(* IEC 61131-3 sources: trust-platform/examples/OSCAT/cleanroom_pressure_strategy_composite/oop/src, 3 files *)

(* ---- Main.st ---- *)
(* Pattern role: IRoomNode is the contract boundary for the Strategy and Composite example. *)
INTERFACE IRoomNode
    PROPERTY ChildCount : INT
    GET
    END_GET
    END_PROPERTY
    PROPERTY PressureError : REAL
    GET
    END_GET
    END_PROPERTY
    PROPERTY AlarmCount : INT
    GET
    END_GET
    END_PROPERTY
    METHOD GetChild : IRoomNode
    VAR_INPUT
        Index : INT;
    END_VAR
    END_METHOD
END_INTERFACE

(* Pattern role: IPressureStrategy is the contract boundary for the Strategy and Composite example. *)
INTERFACE IPressureStrategy
    PROPERTY ModeId : INT
    GET
    END_GET
    END_PROPERTY
    METHOD TargetPressure : REAL
    VAR_INPUT
        BasePressurePa : REAL;
    END_VAR
    END_METHOD
END_INTERFACE

(* Pattern role: NormalPressureStrategy is a concrete implementation in the Strategy and Composite example. *)
FUNCTION_BLOCK NormalPressureStrategy IMPLEMENTS IPressureStrategy
METHOD PUBLIC TargetPressure : REAL
VAR_INPUT
    BasePressurePa : REAL;
END_VAR
TargetPressure := BasePressurePa;
END_METHOD
PUBLIC PROPERTY ModeId : INT
GET
    ModeId := INT#1;
END_GET
END_PROPERTY
END_FUNCTION_BLOCK

(* Pattern role: CleaningPressureStrategy is a concrete implementation in the Strategy and Composite example. *)
FUNCTION_BLOCK CleaningPressureStrategy IMPLEMENTS IPressureStrategy
METHOD PUBLIC TargetPressure : REAL
VAR_INPUT
    BasePressurePa : REAL;
END_VAR
TargetPressure := BasePressurePa + REAL#5.0;
END_METHOD
PUBLIC PROPERTY ModeId : INT
GET
    ModeId := INT#2;
END_GET
END_PROPERTY
END_FUNCTION_BLOCK

(* Pattern role: EmergencyPressureStrategy is a concrete implementation in the Strategy and Composite example. *)
FUNCTION_BLOCK EmergencyPressureStrategy IMPLEMENTS IPressureStrategy
METHOD PUBLIC TargetPressure : REAL
VAR_INPUT
    BasePressurePa : REAL;
END_VAR
TargetPressure := REAL#0.0;
END_METHOD
PUBLIC PROPERTY ModeId : INT
GET
    ModeId := INT#3;
END_GET
END_PROPERTY
END_FUNCTION_BLOCK

(* Pattern role: RoomNode is a concrete implementation in the Strategy and Composite example. *)
FUNCTION_BLOCK RoomNode IMPLEMENTS IRoomNode
VAR
    ErrorValue : REAL;
    AlarmValue : BOOL;
END_VAR
METHOD PUBLIC UpdateRoom
VAR_INPUT
    ActualPressurePa : REAL;
    TargetPressurePa : REAL;
    DoorOpen : BOOL;
END_VAR
ErrorValue := TargetPressurePa - ActualPressurePa;
AlarmValue := (ABS(ErrorValue) > REAL#10.0) OR DoorOpen;
END_METHOD
METHOD PUBLIC GetChild : IRoomNode
VAR_INPUT
    Index : INT;
END_VAR
GetChild := THIS;
END_METHOD
PUBLIC PROPERTY ChildCount : INT
GET
    ChildCount := INT#0;
END_GET
END_PROPERTY
PUBLIC PROPERTY PressureError : REAL
GET
    PressureError := ErrorValue;
END_GET
END_PROPERTY
PUBLIC PROPERTY AlarmCount : INT
GET
    IF AlarmValue THEN AlarmCount := INT#1; ELSE AlarmCount := INT#0; END_IF;
END_GET
END_PROPERTY
END_FUNCTION_BLOCK

(* Pattern role: RoomSuite is a concrete implementation in the Strategy and Composite example. *)
FUNCTION_BLOCK RoomSuite IMPLEMENTS IRoomNode
VAR
    Room1 : RoomNode;
    Room2 : RoomNode;
END_VAR
METHOD PUBLIC UpdateSuite
VAR_INPUT
    Room1Pressure : REAL;
    Room2Pressure : REAL;
    TargetPressure : REAL;
    DoorOpen : BOOL;
END_VAR
Room1.UpdateRoom(ActualPressurePa := Room1Pressure, TargetPressurePa := TargetPressure, DoorOpen := DoorOpen);
Room2.UpdateRoom(ActualPressurePa := Room2Pressure, TargetPressurePa := TargetPressure - REAL#5.0, DoorOpen := FALSE);
END_METHOD
METHOD PUBLIC GetChild : IRoomNode
VAR_INPUT
    Index : INT;
END_VAR
IF Index = INT#1 THEN GetChild := Room1; ELSE GetChild := Room2; END_IF;
END_METHOD
PUBLIC PROPERTY ChildCount : INT
GET
    ChildCount := INT#2;
END_GET
END_PROPERTY
PUBLIC PROPERTY PressureError : REAL
GET
    PressureError := Room1.PressureError + Room2.PressureError;
END_GET
END_PROPERTY
PUBLIC PROPERTY AlarmCount : INT
GET
    AlarmCount := Room1.AlarmCount + Room2.AlarmCount;
END_GET
END_PROPERTY
END_FUNCTION_BLOCK

(* Composition role: PressureCascadeController owns the collaborating objects used by this Strategy and Composite example. *)
FUNCTION_BLOCK PressureCascadeController
VAR
    Normal : NormalPressureStrategy;
    Cleaning : CleaningPressureStrategy;
    Emergency : EmergencyPressureStrategy;
    ActiveStrategy : IPressureStrategy;
    Suite : RoomSuite;
    ActiveModeIdValue : INT;
    SupplyDamperCommandValue : REAL;
END_VAR
METHOD PUBLIC Initialize
ActiveStrategy := Normal;
END_METHOD
METHOD PUBLIC Update : REAL
VAR_INPUT
    ModeRequest : INT;
    Room1Pressure : REAL;
    Room2Pressure : REAL;
    DoorOpen : BOOL;
END_VAR
VAR
    Target : REAL;
END_VAR
IF ModeRequest = INT#3 THEN
    ActiveStrategy := Emergency;
ELSIF ModeRequest = INT#2 THEN
    ActiveStrategy := Cleaning;
ELSE
    ActiveStrategy := Normal;
END_IF;
ActiveModeIdValue := ActiveStrategy.ModeId;
Target := ActiveStrategy.TargetPressure(BasePressurePa := REAL#15.0);
Suite.UpdateSuite(Room1Pressure := Room1Pressure, Room2Pressure := Room2Pressure, TargetPressure := Target, DoorOpen := DoorOpen);
SupplyDamperCommandValue := LIMIT(REAL#0.0, Suite.PressureError * REAL#2.0, REAL#100.0);
Update := SupplyDamperCommandValue;
END_METHOD
PUBLIC PROPERTY ActiveModeId : INT
GET
    ActiveModeId := ActiveModeIdValue;
END_GET
END_PROPERTY
PUBLIC PROPERTY SupplyDamperCommand : REAL
GET
    SupplyDamperCommand := SupplyDamperCommandValue;
END_GET
END_PROPERTY
PUBLIC PROPERTY AlarmCount : INT
GET
    AlarmCount := Suite.AlarmCount;
END_GET
END_PROPERTY
END_FUNCTION_BLOCK

(* Scan role: Main wires the example objects and exposes the PLC call path under test. *)
PROGRAM Main
VAR
    Cascade : PressureCascadeController;
    ModeRequest : INT;
    Room1PressureRaw : INT;
    Room2PressureRaw : INT;
    DoorOpen : BOOL;
    SupplyDamperRaw : INT;
    AlarmOut : BOOL;
END_VAR
Cascade.Initialize();
SupplyDamperRaw := REAL_TO_INT(Cascade.Update(ModeRequest := ModeRequest, Room1Pressure := INT_TO_REAL(Room1PressureRaw), Room2Pressure := INT_TO_REAL(Room2PressureRaw), DoorOpen := DoorOpen));
AlarmOut := Cascade.AlarmCount > INT#0;
END_PROGRAM

(* ---- Configuration.st ---- *)
CONFIGURATION CleanroomPressureStrategyCompositeOopConfiguration
RESOURCE Cpu0 ON PLC
    TASK MainTask (INTERVAL := T#100ms, PRIORITY := 1);
    PROGRAM Cascade WITH MainTask : Main;
END_RESOURCE
VAR_CONFIG
    Cascade.ModeRequest AT %IW0 : INT;
    Cascade.Room1PressureRaw AT %IW2 : INT;
    Cascade.Room2PressureRaw AT %IW4 : INT;
    Cascade.DoorOpen AT %IX0.0 : BOOL;
    Cascade.SupplyDamperRaw AT %QW0 : INT;
    Cascade.AlarmOut AT %QX0.0 : BOOL;
END_VAR
END_CONFIGURATION

(* ---- Tests.st ---- *)
TEST_PROGRAM CleanroomStrategiesChangeTarget
VAR
    Cascade : PressureCascadeController;
    NormalCmd : REAL;
    CleaningCmd : REAL;
END_VAR
Cascade.Initialize();
NormalCmd := Cascade.Update(ModeRequest := INT#1, Room1Pressure := REAL#10.0, Room2Pressure := REAL#5.0, DoorOpen := FALSE);
CleaningCmd := Cascade.Update(ModeRequest := INT#2, Room1Pressure := REAL#10.0, Room2Pressure := REAL#5.0, DoorOpen := FALSE);
ASSERT_TRUE(IN := CleaningCmd > NormalCmd);
ASSERT_EQUAL(EXPECTED := INT#2, ACTUAL := Cascade.ActiveModeId);
END_TEST_PROGRAM

TEST_PROGRAM CleanroomCompositeAggregatesRoomAlarms
VAR
    Cascade : PressureCascadeController;
    Cmd : REAL;
END_VAR
Cascade.Initialize();
Cmd := Cascade.Update(ModeRequest := INT#1, Room1Pressure := REAL#0.0, Room2Pressure := REAL#0.0, DoorOpen := TRUE);
ASSERT_TRUE(IN := Cascade.AlarmCount > INT#0);
END_TEST_PROGRAM

(* Mode-cycling integration test: drives the same Cascade through
   Normal -> Cleaning -> Emergency -> Normal mode requests. Catches
   bugs where the previous strategy's state leaks into the new mode,
   or where ActiveModeId fails to reflect the latest request. *)
TEST_PROGRAM CleanroomCascadeCyclesAllStrategiesOnOneInstance
VAR
    Cascade : PressureCascadeController;
    Cmd : REAL;
END_VAR

Cascade.Initialize();

(* Normal mode *)
Cmd := Cascade.Update(ModeRequest := INT#1, Room1Pressure := REAL#10.0, Room2Pressure := REAL#5.0, DoorOpen := FALSE);
ASSERT_EQUAL(EXPECTED := INT#1, ACTUAL := Cascade.ActiveModeId);

(* Cleaning mode *)
Cmd := Cascade.Update(ModeRequest := INT#2, Room1Pressure := REAL#10.0, Room2Pressure := REAL#5.0, DoorOpen := FALSE);
ASSERT_EQUAL(EXPECTED := INT#2, ACTUAL := Cascade.ActiveModeId);

(* Emergency mode *)
Cmd := Cascade.Update(ModeRequest := INT#3, Room1Pressure := REAL#10.0, Room2Pressure := REAL#5.0, DoorOpen := FALSE);
ASSERT_EQUAL(EXPECTED := INT#3, ACTUAL := Cascade.ActiveModeId);

(* Back to Normal — the strategy slot must reassign cleanly *)
Cmd := Cascade.Update(ModeRequest := INT#1, Room1Pressure := REAL#10.0, Room2Pressure := REAL#5.0, DoorOpen := FALSE);
ASSERT_EQUAL(EXPECTED := INT#1, ACTUAL := Cascade.ActiveModeId);
END_TEST_PROGRAM

(* Strategies in isolation: each FB returns the documented target.
   Catches a future regression where the ModeId getter and the
   TargetPressure delta drift apart. *)
TEST_PROGRAM CleanroomStrategiesInIsolationProduceCorrectTargets
VAR
    Normal : NormalPressureStrategy;
    Cleaning : CleaningPressureStrategy;
    Emergency : EmergencyPressureStrategy;
END_VAR

ASSERT_EQUAL(EXPECTED := INT#1, ACTUAL := Normal.ModeId);
ASSERT_EQUAL(EXPECTED := INT#2, ACTUAL := Cleaning.ModeId);
ASSERT_EQUAL(EXPECTED := INT#3, ACTUAL := Emergency.ModeId);
ASSERT_NEAR(EXPECTED := REAL#15.0, ACTUAL := Normal.TargetPressure(BasePressurePa := REAL#15.0), DELTA := REAL#0.001);
ASSERT_NEAR(EXPECTED := REAL#20.0, ACTUAL := Cleaning.TargetPressure(BasePressurePa := REAL#15.0), DELTA := REAL#0.001);
ASSERT_NEAR(EXPECTED := REAL#0.0, ACTUAL := Emergency.TargetPressure(BasePressurePa := REAL#15.0), DELTA := REAL#0.001);
END_TEST_PROGRAM

(* RoomSuite composite walks both children. ChildCount and AlarmCount
   must aggregate from the two RoomNode children, not be hard-coded
   on the parent. *)
TEST_PROGRAM CleanroomCompositeAggregatesAcrossBothChildren
VAR
    Suite : RoomSuite;
END_VAR

(* Both rooms healthy: zero alarms *)
Suite.UpdateSuite(Room1Pressure := REAL#15.0, Room2Pressure := REAL#10.0, TargetPressure := REAL#15.0, DoorOpen := FALSE);
ASSERT_EQUAL(EXPECTED := INT#2, ACTUAL := Suite.ChildCount);
ASSERT_EQUAL(EXPECTED := INT#0, ACTUAL := Suite.AlarmCount);
(* Room1 fault only: AlarmCount = 1 *)
Suite.UpdateSuite(Room1Pressure := REAL#0.0, Room2Pressure := REAL#10.0, TargetPressure := REAL#15.0, DoorOpen := FALSE);
ASSERT_EQUAL(EXPECTED := INT#1, ACTUAL := Suite.AlarmCount);
(* Both rooms faulted: AlarmCount = 2 *)
Suite.UpdateSuite(Room1Pressure := REAL#0.0, Room2Pressure := REAL#100.0, TargetPressure := REAL#15.0, DoorOpen := FALSE);
ASSERT_EQUAL(EXPECTED := INT#2, ACTUAL := Suite.AlarmCount);
END_TEST_PROGRAM

(* Emergency strategy zeroes the target regardless of base pressure.
   The damper command must respond to the new target on the same scan,
   not lag a cycle. *)
TEST_PROGRAM CleanroomEmergencyDrivesZeroPressureOnSameCycle
VAR
    Cascade : PressureCascadeController;
    Cmd : REAL;
END_VAR

Cascade.Initialize();
(* Establish baseline at Normal mode *)
Cmd := Cascade.Update(ModeRequest := INT#1, Room1Pressure := REAL#15.0, Room2Pressure := REAL#10.0, DoorOpen := FALSE);
(* Switch to Emergency: target = 0; Room1 above target by 15 Pa, Room2 by 15 Pa *)
Cmd := Cascade.Update(ModeRequest := INT#3, Room1Pressure := REAL#15.0, Room2Pressure := REAL#10.0, DoorOpen := FALSE);
ASSERT_EQUAL(EXPECTED := INT#3, ACTUAL := Cascade.ActiveModeId);
(* PressureError = (0 - 15) + ((0 - 5) - 10) = -30; clamped to 0 *)
ASSERT_NEAR(EXPECTED := REAL#0.0, ACTUAL := Cmd, DELTA := REAL#0.001);
END_TEST_PROGRAM

(* Damper command saturation: a far-from-target pressure clamps to 100,
   it does not overshoot. The LIMIT call inside Update is the gate. *)
TEST_PROGRAM CleanroomDamperCommandSaturatesAtHighEnd
VAR
    Cascade : PressureCascadeController;
    Cmd : REAL;
END_VAR

Cascade.Initialize();
(* Normal mode target = 15; both rooms read 0 -> error sum = 25, *2 = 50 *)
Cmd := Cascade.Update(ModeRequest := INT#1, Room1Pressure := REAL#0.0, Room2Pressure := REAL#0.0, DoorOpen := FALSE);
ASSERT_TRUE(IN := Cmd <= REAL#100.0);
(* Cleaning mode target = 20; both rooms read 0 -> error sum = 35, *2 = 70 *)
Cmd := Cascade.Update(ModeRequest := INT#2, Room1Pressure := REAL#0.0, Room2Pressure := REAL#0.0, DoorOpen := FALSE);
ASSERT_TRUE(IN := Cmd <= REAL#100.0);
ASSERT_TRUE(IN := Cmd >= REAL#0.0);
END_TEST_PROGRAM

(* DoorOpen on a healthy suite still triggers alarm in Room1 only.
   Room2 is intentionally not exposed to door state in this demo. *)
TEST_PROGRAM CleanroomDoorOpenAlarmsRoom1Only
VAR
    Cascade : PressureCascadeController;
    Cmd : REAL;
END_VAR

Cascade.Initialize();
(* Normal mode, both rooms exactly at target, door open *)
Cmd := Cascade.Update(ModeRequest := INT#1, Room1Pressure := REAL#15.0, Room2Pressure := REAL#10.0, DoorOpen := TRUE);
ASSERT_EQUAL(EXPECTED := INT#1, ACTUAL := Cascade.AlarmCount);
(* Same pressures, door closed: no alarm *)
Cmd := Cascade.Update(ModeRequest := INT#1, Room1Pressure := REAL#15.0, Room2Pressure := REAL#10.0, DoorOpen := FALSE);
ASSERT_EQUAL(EXPECTED := INT#0, ACTUAL := Cascade.AlarmCount);
END_TEST_PROGRAM
